// TIA Portal V21 export
// export: Created 2026-11-08T21:21:44.3073789Z, ExportSetting WithDefaults, DisplayName Totally Integrated Automation Portal, DisplayVersion V21 Update 3, DisplayName STEP 7 Professional, DisplayVersion V21 Update 3, DisplayName STEP 7 Safety, DisplayVersion V21, DisplayName Tech WebApplication, DisplayVersion V21, DisplayName WinCC Basic/Comfort/Advanced, DisplayVersion V21 Update 3, DisplayName WinCC Unified, DisplayVersion V21 Update 3
FUNCTION "FC_StlPar" : Void   // FC3, STL
{ S7_Optimized_Access := 'TRUE' }
VERSION : 0.1
// stored: AutoNumber true, UDAEnableTagReadback false
   VAR_INPUT
      x : Int;
      y : Int;
   END_VAR
   VAR_OUTPUT
      q : Bool;
      r : Int;
   END_VAR
BEGIN

NETWORK
TITLE = 
      L     #x;
      L     #y;
      +I;
      T     #r;
      >I;
      =     #q;
END_FUNCTION
